Fanuc KAREL source: kb00019.compact.KL

PROGRAM KB00019
%STACKSIZE=65535
%PRIORITY=65535
%NOLOCKGROUP
%ENVIRONMENT FDEV
VAR
P1 : STRING[80]
P2 : INTEGER
BEGIN
P1='A'
P2=1
CHECK_NAME(P1,P2)
END KB00019
